FUNCTION_BLOCK GATE_CYCLE (* Migrated from IEC 61131-3 ST *)
  (* Standard: 61499-2 *)
  (* Version 1.0, 2026-11-06, st2fb *)
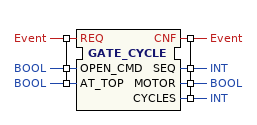
  EVENT_INPUT
    REQ WITH OPEN_CMD, AT_TOP;
  END_EVENT
  EVENT_OUTPUT
    CNF WITH SEQ, MOTOR, CYCLES;
  END_EVENT
  VAR_INPUT
    OPEN_CMD : BOOL;
    AT_TOP : BOOL;
  END_VAR
  VAR_OUTPUT
    SEQ : INT;
    MOTOR : BOOL;
    CYCLES : INT;
  END_VAR
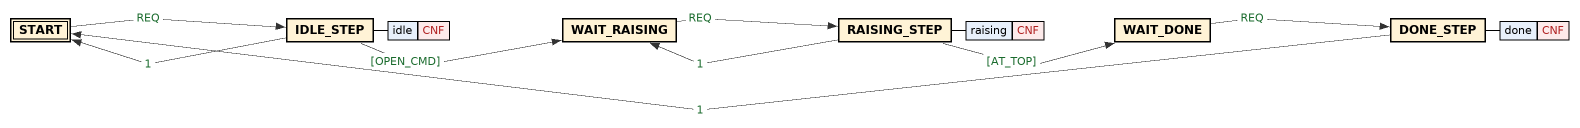
  EC_STATES
    START;
    IDLE_STEP : idle -> CNF;
    WAIT_RAISING;
    RAISING_STEP : raising -> CNF;
    WAIT_DONE;
    DONE_STEP : done -> CNF;
  END_STATES
  EC_TRANSITIONS
    START TO IDLE_STEP := REQ;
    IDLE_STEP TO WAIT_RAISING := [OPEN_CMD];
    IDLE_STEP TO START := 1;
    WAIT_RAISING TO RAISING_STEP := REQ;
    RAISING_STEP TO WAIT_DONE := [AT_TOP];
    RAISING_STEP TO WAIT_RAISING := 1;
    WAIT_DONE TO DONE_STEP := REQ;
    DONE_STEP TO START := 1;
  END_TRANSITIONS
  ALGORITHM idle IN ST:
MOTOR := FALSE;
IF OPEN_CMD THEN
  SEQ := 1;
END_IF;
  END_ALGORITHM
  ALGORITHM raising IN ST:
MOTOR := TRUE;
IF AT_TOP THEN
  SEQ := 2;
END_IF;
  END_ALGORITHM
  ALGORITHM done IN ST:
MOTOR := FALSE;
CYCLES := CYCLES + 1;
SEQ := 0;
  END_ALGORITHM
END_FUNCTION_BLOCK
